Fanuc KAREL source: KB00098.KL

PROGRAM KB00098
%NOLOCKGROUP
%ENVIRONMENT TIM
VAR
  P1: INTEGER
  P2: INTEGER
BEGIN
  P1 = 1
  P2 = 1
  GET_USEC_SUB(P1, P2)
END KB00098
